FUNCTION "Mode_Change_F"   // FC 2, author

VAR_INPUT
   Mode : UInt;
END_VAR

VAR_TEMP
   i : UInt;
   j : UInt;
END_VAR

   // RETURN : Void
BEGIN
// REGION Change all devices
//     "Control_DB".ECnv_Control.Instruction.Mode_Change := #Mode;
//     "Control_DB".VTD_Control.Instruction.Mode_Change := #Mode;

//     FOR #i := "Settings_DB".VTD_Settings.Lowest_Level TO "Settings_DB".VTD_Settings.Highest_Level DO
//         "Control_DB".LCnv_Control.Cnv_Level_Control[#i].Cnv1_Control.Instruction.Mode_Change := #Mode;
//         "Control_DB".LCnv_Control.Cnv_Level_Control[#i].Cnv2_Control.Instruction.Mode_Change := #Mode;
//     END_FOR;
// END_REGION



END_FUNCTION